PROGRAM main
  VAR
    S1 AT %IX0.0  : BOOL; (* marcha, NA *)
    S2 AT %IX0.1  : BOOL; (* paro, NC: TRUE sin pulsar *)
    KM1 AT %QX0.0 : BOOL; (* motor *)
    H1 AT %QX0.1  : BOOL; (* mantenimiento *)
    T_SEG         : TON;
    PULSO         : BOOL; (* TRUE una vuelta por segundo de marcha *)
    SEGUNDOS      : INT; (* horómetro: segundos de marcha *)
    HAY_TIEMPO    : BOOL; (* SEGUNDOS < 20 *)
  END_VAR
  VAR  (* added by the conversion: wires and edge detectors of the diagram *)
    _LT1_OUT : BOOL;
    _OR6_OUT : BOOL;
    _AND5_OUT : BOOL;
    _NOT15_OUT : BOOL;
    _AND13_OUT : BOOL;
    _ADD22_OUT : INT;
    _SEL19_OUT : INT;
    _GE26_OUT : BOOL;
  END_VAR

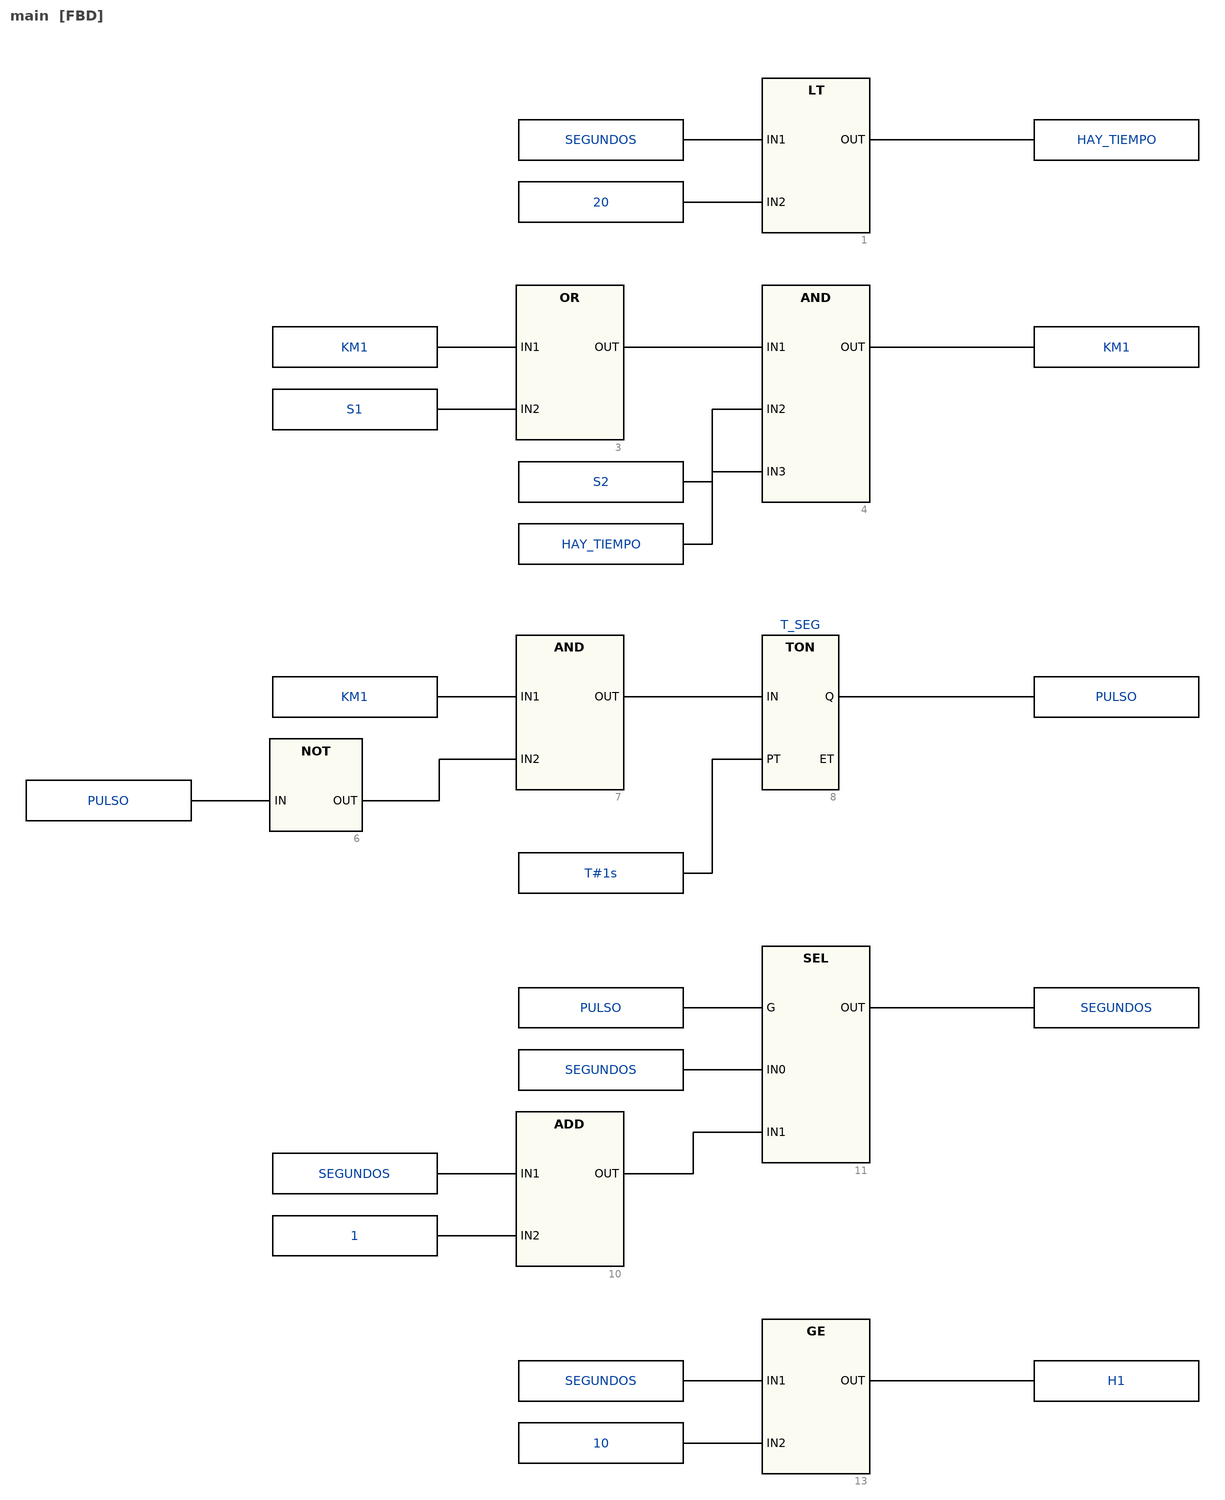
(* FBD diagram, written out as Structured Text *)
_LT1_OUT := SEGUNDOS < 20;
HAY_TIEMPO := _LT1_OUT;
_OR6_OUT := KM1 OR S1;
_AND5_OUT := _OR6_OUT AND S2 AND HAY_TIEMPO;
KM1 := _AND5_OUT;
_NOT15_OUT := NOT PULSO;
_AND13_OUT := KM1 AND _NOT15_OUT;
T_SEG(IN := _AND13_OUT, PT := T#1s);
PULSO := T_SEG.Q;
_ADD22_OUT := SEGUNDOS + 1;
_SEL19_OUT := SEL(PULSO, SEGUNDOS, _ADD22_OUT);
SEGUNDOS := _SEL19_OUT;
_GE26_OUT := SEGUNDOS >= 10;
H1 := _GE26_OUT;
END_PROGRAM
